TYPE "DT_MEASUREMENT_SYSTEM_GENERATOR_MEASUREMENT"
VERSION : 0.1
   STRUCT
      I_1 { S7_SetPoint := 'False'} : "DT_MEASUREMENT_SOLO" := ((), (), FALSE, 1, 0, 48, 32000, 32000, 32000, 0, 0, 0, 0, 0, 0, 0, 0, 0, 0, 0, 0, 0, 0.0, '');
      I_2 { S7_SetPoint := 'False'} : "DT_MEASUREMENT_SOLO" := ((), (), FALSE, 1, 0, 49, 32000, 32000, 32000, 0, 0, 0, 0, 0, 0, 0, 0, 0, 0, 0, 0, 0, 0.0, '');
      I_3 { S7_SetPoint := 'False'} : "DT_MEASUREMENT_SOLO" := ((), (), FALSE, 1, 0, 50, 32000, 32000, 32000, 0, 0, 0, 0, 0, 0, 0, 0, 0, 0, 0, 0, 0, 0.0, '');
      I { S7_SetPoint := 'False'} : "DT_MEASUREMENT_SOLO" := ((), (), FALSE, 1, 0, 51, 32000, 32000, 32000, 0, 0, 0, 0, 0, 0, 0, 0, 0, 0, 0, 0, 0, 0.0, '');
      U12 { S7_SetPoint := 'False'} : "DT_MEASUREMENT_SOLO" := ((), (), FALSE, 1, 0, 52, 32000, 32000, 32000, 0, 0, 0, 0, 0, 0, 0, 0, 0, 0, 0, 0, 0, 0.0, '');
      U13 { S7_SetPoint := 'False'} : "DT_MEASUREMENT_SOLO" := ((), (), FALSE, 1, 0, 53, 32000, 32000, 32000, 0, 0, 0, 0, 0, 0, 0, 0, 0, 0, 0, 0, 0, 0.0, '');
      U23 { S7_SetPoint := 'False'} : "DT_MEASUREMENT_SOLO" := ((), (), FALSE, 1, 0, 54, 32000, 32000, 32000, 0, 0, 0, 0, 0, 0, 0, 0, 0, 0, 0, 0, 0, 0.0, '');
      U_LL { S7_SetPoint := 'False'} : "DT_MEASUREMENT_SOLO" := ((), (), FALSE, 1, 0, 55, 32000, 32000, 32000, 0, 0, 0, 0, 0, 0, 0, 0, 0, 0, 0, 0, 0, 0.0, '');
      U1 { S7_SetPoint := 'False'} : "DT_MEASUREMENT_SOLO" := ((), (), FALSE, 1, 0, 56, 32000, 32000, 32000, 0, 0, 0, 0, 0, 0, 0, 0, 0, 0, 0, 0, 0, 0.0, '');
      U2 { S7_SetPoint := 'False'} : "DT_MEASUREMENT_SOLO" := ((), (), FALSE, 1, 0, 57, 32000, 32000, 32000, 0, 0, 0, 0, 0, 0, 0, 0, 0, 0, 0, 0, 0, 0.0, '');
      U3 { S7_SetPoint := 'False'} : "DT_MEASUREMENT_SOLO" := ((), (), FALSE, 1, 0, 58, 32000, 32000, 32000, 0, 0, 0, 0, 0, 0, 0, 0, 0, 0, 0, 0, 0, 0.0, '');
      f { S7_SetPoint := 'False'} : "DT_MEASUREMENT_SOLO" := ((), (), FALSE, 1, 0, 59, 32000, 32000, 32000, 0, 0, 0, 0, 0, 0, 0, 0, 0, 0, 0, 0, 0, 0.0, '');
      PF { S7_SetPoint := 'False'} : "DT_MEASUREMENT_SOLO" := ((), (), FALSE, 1, 0, 60, 32000, 32000, 32000, 0, 0, 0, 0, 0, 0, 0, 0, 0, 0, 0, 0, 0, 0.0, '');
      P { S7_SetPoint := 'False'} : "DT_MEASUREMENT_SOLO" := ((), (), FALSE, 1, 0, 61, 32000, 32000, 32000, 0, 0, 0, 0, 0, 0, 0, 0, 0, 0, 0, 0, 0, 0.0, '');
      Q { S7_SetPoint := 'False'} : "DT_MEASUREMENT_SOLO" := ((), (), FALSE, 1, 0, 62, 32000, 32000, 32000, 0, 0, 0, 0, 0, 0, 0, 0, 0, 0, 0, 0, 0, 0.0, '');
      S { S7_SetPoint := 'False'} : "DT_MEASUREMENT_SOLO" := ((), (), FALSE, 1, 0, 63, 32000, 32000, 32000, 0, 0, 0, 0, 0, 0, 0, 0, 0, 0, 0, 0, 0, 0.0, '');
      E_ACT_IMP { S7_SetPoint := 'False'} : "DT_MEASUREMENT_SOLO" := ((), (), FALSE, 1, 0, 64, 32000, 32000, 32000, 0, 0, 0, 0, 0, 0, 0, 0, 0, 0, 0, 0, 0, 0.0, '');
      E_ACT_EXP { S7_SetPoint := 'False'} : "DT_MEASUREMENT_SOLO" := ((), (), FALSE, 1, 0, 65, 32000, 32000, 32000, 0, 0, 0, 0, 0, 0, 0, 0, 0, 0, 0, 0, 0, 0.0, '');
      E_RACT_IMP { S7_SetPoint := 'False'} : "DT_MEASUREMENT_SOLO" := ((), (), FALSE, 1, 0, 66, 32000, 32000, 32000, 0, 0, 0, 0, 0, 0, 0, 0, 0, 0, 0, 0, 0, 0.0, '');
      E_RACT_EXP { S7_SetPoint := 'False'} : "DT_MEASUREMENT_SOLO" := ((), (), FALSE, 1, 0, 67, 32000, 32000, 32000, 0, 0, 0, 0, 0, 0, 0, 0, 0, 0, 0, 0, 0, 0.0, '');
      MEAS_20 { S7_SetPoint := 'False'} : "DT_MEASUREMENT_SOLO" := ((), (), FALSE, 1, 0, 68, 32000, 32000, 32000, 0, 0, 0, 0, 0, 0, 0, 0, 0, 0, 0, 0, 0, 0.0, '');
      MEAS_21 { S7_SetPoint := 'False'} : "DT_MEASUREMENT_SOLO" := ((), (), FALSE, 1, 0, 69, 32000, 32000, 32000, 0, 0, 0, 0, 0, 0, 0, 0, 0, 0, 0, 0, 0, 0.0, '');
      MEAS_22 { S7_SetPoint := 'False'} : "DT_MEASUREMENT_SOLO" := ((), (), FALSE, 1, 0, 70, 32000, 32000, 32000, 0, 0, 0, 0, 0, 0, 0, 0, 0, 0, 0, 0, 0, 0.0, '');
      MEAS_23 { S7_SetPoint := 'False'} : "DT_MEASUREMENT_SOLO" := ((), (), FALSE, 1, 0, 71, 32000, 32000, 32000, 0, 0, 0, 0, 0, 0, 0, 0, 0, 0, 0, 0, 0, 0.0, '');
   END_STRUCT;

END_TYPE

